FUNCTION_BLOCK T_E_text_EtherCAT EXTENDS T_E_text_Common
VAR
END_VAR

PROPERTY allDevicesOk : KOSTAL_AF2024_Core_Text.ST_E_Text
GET
allDevicesOk.Number:= 11;
END_GET
END_PROPERTY

PROPERTY device_0_isInState_1 : KOSTAL_AF2024_Core_Text.ST_E_Text
GET
device_0_isInState_1.Number:= 10;
END_GET
END_PROPERTY

PROPERTY name : KOSTAL_AF2024_Core_Text.ST_E_Text
GET
name.Number:= 2;
END_GET
END_PROPERTY

END_FUNCTION_BLOCK

(* stored: Version 1.1.0.1, ProductVersion 3.1.4024.12
   POU T_E_text_EtherCAT: Id {cd64bb43-835f-4e86-984e-5d77e1ca43e3}, SpecialFunc None
   Property allDevicesOk: Id {1d235980-4095-4c20-b1bd-73314e95f820}
   Get Get: Id {e84e57ce-ced0-4747-8eb8-ee1d39e5628f}
   Property device_0_isInState_1: Id {7105d90c-0836-4173-aeb3-65d99943006a}
   Get Get: Id {62ff15f1-76ee-4745-a4df-9ba4ef4f93b8}
   Property name: Id {a4f69d73-a869-4901-a280-39e2fac8e5f3}
   Get Get: Id {8a0472f2-2aea-4d79-9be2-22ee1dc92ad5} *)
